// TIA Portal V19 export
// export: Created 2026-10-15T09:44:24.9895988Z, ExportSetting WithDefaults, DisplayName Totally Integrated Automation Portal, DisplayVersion V19, DisplayName TIA Portal Openness, DisplayVersion V19, DisplayName TIA Portal Version Control Interface, DisplayVersion V19, DisplayName STEP 7 Professional, DisplayVersion V19, DisplayName STEP 7 Safety, DisplayVersion V19, DisplayName WinCC Basic/Comfort/Advanced, DisplayVersion V19, DisplayName WinCC Unified, DisplayVersion V19
FUNCTION "ROLL_PB50" : Void   // FC33, SCL
{ S7_Optimized_Access := 'TRUE' }
VERSION : 0.1
// stored: AutoNumber true, IsIECCheckEnabled false, SetENOAutomatically false, UDAEnableTagReadback false
   VAR_TEMP
      r : Bool;
      a1 : Word;
      a2 : Word;
      activeDataBlock : Int;
      comparisonResults : Array[0..0] of Bool;
   END_VAR
BEGIN

   #r := FALSE;
   #a1 := W#16#0000;
   #a2 := W#16#0000;
   #activeDataBlock := 0;
   // PB50, STEP 5 network 1
   #activeDataBlock := 15;
   // PB50, STEP 5 network 2
   #r := "ROLL_State".M[0, 1];
   IF #r THEN
       "ROLL_State".M[0, 2] := FALSE;
   END_IF;
   // PB50, STEP 5 network 3
   #a2 := #a1;
   #a1 := W#16#2008;
   #r := ((NOT "ROLL_State".M[0, 1]) AND "ROLL_IO".Input[3, 0]);
   "ROLL_TimerOp"(Number := 11,
                  Operation := 0,
                  Signal := #r,
                  Preset := #a1);
   // PB50, STEP 5 network 4
   #a2 := #a1;
   #a1 := W#16#1020;
   #r := "ROLL_State".M[29, 0];
   "ROLL_TimerOp"(Number := 13,
                  Operation := 0,
                  Signal := #r,
                  Preset := #a1);
   // PB50, STEP 5 network 5
   RETURN;
END_FUNCTION
